{attribute 'qualified_only'}
VAR_GLOBAL
	TorqueM1_Act AT %I* : LREAL;
	TorqueM2_Act AT %I* : LREAL;
	TorqueM3_Act AT %I* : LREAL;
	TorqueM33_Act : LREAL;
END_VAR

(* stored: Version 1.1.0.1, ProductVersion 3.1.4024.15
   GVL GVL_Torque: Id {97919b58-756f-46a0-a20b-a3771fa2b570} *)
